Fanuc KAREL source: kc00010.KL

-- PROVISIONAL review KL for V770-1; original PC SHA256 de78efe1a113818548b5c04ccc4303729049700b82aa5125b15e5f24e711ae51
-- Incomplete behavior may be omitted. Consult companion uncertainty JSON. Do not deploy.
PROGRAM KC00010
%NOLOCKGROUP
BEGIN
  -- UNRESOLVED_PC offsets 5-27; opcodes 27,22,1C,31,23
  -- UNRESOLVED_PC offsets 32-36; opcodes 7F
END KC00010
